// TIA Portal V20 export
// export: Created 2026-10-11T05:28:39.8367123Z, ExportSetting WithDefaults, DisplayName Totally Integrated Automation Portal, DisplayVersion V20, DisplayName TIA Portal Openness, DisplayVersion V20, DisplayName TIA Portal Teamcenter Gateway, DisplayVersion V20, DisplayName TIA Portal Version Control Interface, DisplayVersion V20, DisplayName SINAMICS Startdrive Advanced, DisplayVersion V20 SP1 Update 2, DisplayName SINAMICS Startdrive G110M, G120, G120C, G120D, G120P, G115D, DisplayVersion V20 SP1 Update 2, DisplayName SINAMICS Startdrive G130, G150, S120, S150, SINAMICS MV, G220, S200, S210, DisplayVersion V20 SP1 Update 2, DisplayName STEP 7 Professional, DisplayVersion V20, DisplayName STEP 7 Safety, DisplayVersion V20, DisplayName WinCC Basic/Comfort/Advanced, DisplayVersion V20, DisplayName WinCC Professional, DisplayVersion V20, DisplayName WinCC Unified, DisplayVersion V20
FUNCTION "FRK_ConfigAppend" : Void   // FC22, SCL
{ S7_Optimized_Access := 'TRUE' }
VERSION : 0.1
// stored: AutoNumber true, IsIECCheckEnabled false, SetENOAutomatically false, UDAEnableTagReadback false
   VAR_INPUT
      Scope : String;
      Item : String;
      ValueText : WString;
      ValueType : DInt;
      ReadLevel : DInt;
      Readable : Bool;
   END_VAR
   VAR_IN_OUT
      Cursor : "FRK_ConfigCursor";
      Page : "ST_ConfigPage";
   END_VAR
   VAR_TEMP
      Slot : DInt;
   END_VAR
BEGIN

   #Slot := #Cursor.Position - #Cursor.First;
   #Cursor.Position := #Cursor.Position + 1;
   IF #Slot < 0 OR #Slot >= 16 THEN
       RETURN;
   END_IF;
   #Slot := #Slot + 1;
   #Page.Entries[#Slot].Scope := STRING_TO_WSTRING(#Scope);
   #Page.Entries[#Slot].Item := STRING_TO_WSTRING(#Item);
   #Page.Entries[#Slot].ValueType := #ValueType;
   #Page.Entries[#Slot].ReadLevel := #ReadLevel;
   #Page.Entries[#Slot].Readable := #Readable;
   IF #Readable THEN
       #Page.Entries[#Slot].ValueText := #ValueText;
   END_IF;
   #Page.EntryCount := DINT_TO_INT(#Slot);
END_FUNCTION
